FUNCTION_BLOCK FB_Spanner
VAR_INPUT
END_VAR
VAR_OUTPUT
END_VAR
VAR
END_VAR

GVL_IO.xVentilSpannerAS := GVL_IO.xZylinderEinlaufBereit;
GVL_IO.xVentilSpannerGS := NOT GVL_IO.xZylinderEinlaufBereit;
GVL_IO.xSpannerBereit := GVL_IO.xZylinderSpannerAS;

END_FUNCTION_BLOCK

(* stored: Version 1.1.0.1
   POU FB_Spanner: Id {48f5b05a-5920-427c-854a-9de49296cf9a}, SpecialFunc None *)
